// TIA Portal V21 export
// export: Created 2026-11-10T19:11:36.9230349Z, ExportSetting WithDefaults, DisplayName Totally Integrated Automation Portal, DisplayVersion V21 Update 3, DisplayName STEP 7 Professional, DisplayVersion V21 Update 3, DisplayName STEP 7 Safety, DisplayVersion V21, DisplayName Tech WebApplication, DisplayVersion V21, DisplayName WinCC Basic/Comfort/Advanced, DisplayVersion V21 Update 3, DisplayName WinCC Unified, DisplayVersion V21 Update 3
DATA_BLOCK "DB_DRUM"   // DB22
// stored: AutoNumber true, DBAccessibleFromOPCUA true, DBAccessibleFromWebserver true, InstanceOfName DRUM, OfSystemLibElement DRUM, OfSystemLibVersion 2.6
"DRUM"
   // VAR_INPUT
   //    RESET : Bool;
   //    JOG : Bool;
   //    DRUM_EN : Bool;
   //    LST_STEP : Byte;
   //    EVENT1 : Bool;
   //    EVENT2 : Bool;
   //    EVENT3 : Bool;
   //    EVENT4 : Bool;
   //    EVENT5 : Bool;
   //    EVENT6 : Bool;
   //    EVENT7 : Bool;
   //    EVENT8 : Bool;
   //    EVENT9 : Bool;
   //    EVENT10 : Bool;
   //    EVENT11 : Bool;
   //    EVENT12 : Bool;
   //    EVENT13 : Bool;
   //    EVENT14 : Bool;
   //    EVENT15 : Bool;
   //    EVENT16 : Bool;
   // END_VAR
   // VAR_OUTPUT
   //    OUT1 : Bool;
   //    OUT2 : Bool;
   //    OUT3 : Bool;
   //    OUT4 : Bool;
   //    OUT5 : Bool;
   //    OUT6 : Bool;
   //    OUT7 : Bool;
   //    OUT8 : Bool;
   //    OUT9 : Bool;
   //    OUT10 : Bool;
   //    OUT11 : Bool;
   //    OUT12 : Bool;
   //    OUT13 : Bool;
   //    OUT14 : Bool;
   //    OUT15 : Bool;
   //    OUT16 : Bool;
   //    Q : Bool;
   //    OUT_WORD : Word;
   //    ERR_CODE : Word;
   // END_VAR
   // VAR
   //    JOG_HIS : Bool;
   //    EOD : Bool;
   //    DSP : Byte;
   //    DSC : Byte;
   //    DCC : DWord;
   //    DTBP : Word;
   //    PrevTime : Time;
   //    S_PRESET : Array[1..16] of Word;
   //    OUT_VAL : Array[1..16, 0..15] of Bool;
   //    S_MASK : Array[1..16, 0..15] of Bool;
   // END_VAR
BEGIN
END_DATA_BLOCK
